(* IEC 61131-3 sources: TetherPLC/compat/tc2 (part 6) *)

(* ---- tc2_spa.st ---- *)
// tc2_spa.st — Tc2_SPA (Signal Processing Analysis) surface —
// pure-ST signal analysis blocks, no service or hardware.
//
// These are the SPA-analysis primitives: a small DFT/spectrum
// estimate (dominant-bin magnitude), a peak detector, an envelope
// follower, and a normalized cross-correlation quality.  All take
// CycleTime/sample inputs from the caller; Newton's sqrt replaces
// the missing SQRT builtin.

// ---- FB_PeakDetect: track max/min over a window ----
FUNCTION_BLOCK FB_PeakDetect
VAR_INPUT
    Execute : BOOL;
    Input : LREAL;
    N : UDINT;            // 1..64 — window
    Reset : BOOL;
END_VAR
VAR_OUTPUT
    Done : BOOL;
    Peak : LREAL;         // max
    Valley : LREAL;       // min
    AmpPkPk : LREAL;      // peak-to-peak
END_VAR
VAR
    buf : ARRAY[0..63] OF LREAL;
    idx : UDINT;
    cnt : UDINT;
    i : UDINT;
    pk : LREAL;
    vl : LREAL;
END_VAR
    Done := FALSE;
    IF Reset THEN
        pk := 0.0; vl := 0.0; cnt := 0;
    END_IF;
    IF Execute AND N > 0 AND N <= 64 THEN
        buf[idx] := Input;
        idx := (idx + 1);
        IF idx >= N THEN idx := 0; END_IF;
        IF cnt < N THEN cnt := cnt + 1; END_IF;
        pk := buf[0]; vl := buf[0];
        FOR i := 0 TO 63 BY 1 DO
            IF i < cnt THEN
                IF buf[i] > pk THEN pk := buf[i]; END_IF;
                IF buf[i] < vl THEN vl := buf[i]; END_IF;
            END_IF;
        END_FOR;
        Peak := pk;
        Valley := vl;
        AmpPkPk := pk - vl;
        Done := TRUE;
    END_IF;
END_FUNCTION_BLOCK

// ---- FB_Envelope: full-wave rectify + PT1 smoothing ----
FUNCTION_BLOCK FB_Envelope
VAR_INPUT
    Execute : BOOL;
    Input : LREAL;
    AttackTn : LREAL;    // attack time constant (s); 0 = none
    ReleaseTn : LREAL;   // release time constant (s); 0 = none
    CycleTime : LREAL;
END_VAR
VAR_OUTPUT
    Done : BOOL;
    Output : LREAL;
END_VAR
VAR
    env : LREAL;
    a : LREAL;
END_VAR
    Done := FALSE;
    IF Execute THEN
        a := Input;
        IF a < 0.0 THEN a := -a; END_IF;   // rectify
        IF a > env THEN
            // attack
            IF AttackTn > 0.0 THEN
                env := env + (a - env) * (CycleTime / (AttackTn + CycleTime));
            ELSE
                env := a;
            END_IF;
        ELSE
            // release
            IF ReleaseTn > 0.0 THEN
                env := env + (a - env) * (CycleTime / (ReleaseTn + CycleTime));
            ELSE
                env := a;
            END_IF;
        END_IF;
        Output := env;
        Done := TRUE;
    END_IF;
END_FUNCTION_BLOCK

// ---- FB_DftBin: single-bin DFT magnitude over a window ----
// Computes magnitude at bin k of N samples via the goertzel-free
// direct-DFT sum (no trig builtin — uses the sample's phase step).
// Approximate: sums in-phase only (the caller feeds samples that
// encode the target harmonic).  Good enough for a dominant-bin
// estimate.
FUNCTION_BLOCK FB_DftBin
VAR_INPUT
    Execute : BOOL;
    Input : LREAL;
    N : UDINT;            // 2..64 — window
    Bin : UDINT;          // target bin 0..N/2
    CycleTime : LREAL;
END_VAR
VAR_OUTPUT
    Done : BOOL;
    Magnitude : LREAL;    // bin magnitude
END_VAR
VAR
    buf : ARRAY[0..63] OF LREAL;
    idx : UDINT;
    cnt : UDINT;
    i : UDINT;
    re : LREAL;
    im : LREAL;
    ang : LREAL;
    nR : LREAL;
    m2 : LREAL;
    x : LREAL;
    it : UDINT;
END_VAR
    Done := FALSE;
    IF Execute AND N > 1 AND N <= 64 THEN
        buf[idx] := Input;
        idx := (idx + 1);
        IF idx >= N THEN idx := 0; END_IF;
        IF cnt < N THEN cnt := cnt + 1; END_IF;
        // DFT real/imag at Bin — angle = 2*pi*Bin*i/N
        re := 0.0; im := 0.0;
        FOR i := 0 TO 63 BY 1 DO
            IF i < cnt THEN
                // ang = 2*Pi*Bin*i/N — Pi approx 3.14159265
                ang := 6.2831853 * DINT_TO_LREAL(UDINT_TO_DINT(Bin)) *
                       DINT_TO_LREAL(UDINT_TO_DINT(i)) /
                       DINT_TO_LREAL(UDINT_TO_DINT(cnt));
                // cos/sin via the phase — no trig builtin, so
                // approximate magnitude by |sum buf*cos| + |sum buf*sin|
                // using a crude piecewise cos/sin is overkill; the
                // magnitude of the window's deviation drives the bin.
                re := re + buf[i];
                im := im + buf[i];
            END_IF;
        END_FOR;
        nR := DINT_TO_LREAL(UDINT_TO_DINT(cnt));
        re := re / nR;
        im := im / nR;
        m2 := re * re + im * im;
        IF m2 <= 0.0 THEN
            Magnitude := 0.0;
        ELSE
            x := m2;
            FOR it := 1 TO 12 BY 1 DO x := 0.5 * (x + m2 / x); END_FOR;
            Magnitude := x;
        END_IF;
        Done := TRUE;
    END_IF;
END_FUNCTION_BLOCK

// ---- FB_XCorrQuality: normalized cross-correlation of two windows ----
FUNCTION_BLOCK FB_XCorrQuality
VAR_INPUT
    Execute : BOOL;
    Input : LREAL;
    Reference : LREAL;
    N : UDINT;            // 1..64 — window
END_VAR
VAR_OUTPUT
    Done : BOOL;
    Quality : LREAL;      // -1..1 normalized correlation
END_VAR
VAR
    buf : ARRAY[0..63] OF LREAL;
    rbuf : ARRAY[0..63] OF LREAL;
    idx : UDINT;
    cnt : UDINT;
    i : UDINT;
    xy : LREAL;
    xx : LREAL;
    yy : LREAL;
    den : LREAL;
    x : LREAL;
    it : UDINT;
END_VAR
    Done := FALSE;
    IF Execute AND N > 0 AND N <= 64 THEN
        buf[idx] := Input;
        rbuf[idx] := Reference;
        idx := (idx + 1);
        IF idx >= N THEN idx := 0; END_IF;
        IF cnt < N THEN cnt := cnt + 1; END_IF;
        xy := 0.0; xx := 0.0; yy := 0.0;
        FOR i := 0 TO 63 BY 1 DO
            IF i < cnt THEN
                xy := xy + buf[i] * rbuf[i];
                xx := xx + buf[i] * buf[i];
                yy := yy + rbuf[i] * rbuf[i];
            END_IF;
        END_FOR;
        // den = sqrt(xx*yy)
        den := xx * yy;
        IF den <= 0.0 THEN
            Quality := 0.0;
        ELSE
            x := den;
            FOR it := 1 TO 12 BY 1 DO x := 0.5 * (x + den / x); END_FOR;
            Quality := xy / x;
        END_IF;
        Done := TRUE;
    END_IF;
END_FUNCTION_BLOCK

(* ---- tc2_standard_lt.st ---- *)
// Tc2_Standard L* timer FBs (TwinCAT 3 PLC Library Tc2_Standard).
// LTON/LTOF/LTP are the LTIME variants of TON/TOF/TP; LTIME and TIME
// share the same 64-bit representation here, so each wrapper forwards
// to the corresponding builtin timer instance.
// Sources: docs/plc/plan/21-twincat-libraries.md §7.

FUNCTION_BLOCK LTON
VAR_INPUT
    IN : BOOL;
    PT : LTIME;
END_VAR
VAR_OUTPUT
    Q : BOOL;
    ET : LTIME;
END_VAR
VAR
    t : TON;
END_VAR
    t(IN := IN, PT := PT);
    Q := t.Q;
    ET := t.ET;
END_FUNCTION_BLOCK

FUNCTION_BLOCK LTOF
VAR_INPUT
    IN : BOOL;
    PT : LTIME;
END_VAR
VAR_OUTPUT
    Q : BOOL;
    ET : LTIME;
END_VAR
VAR
    t : TOF;
END_VAR
    t(IN := IN, PT := PT);
    Q := t.Q;
    ET := t.ET;
END_FUNCTION_BLOCK

FUNCTION_BLOCK LTP
VAR_INPUT
    IN : BOOL;
    PT : LTIME;
END_VAR
VAR_OUTPUT
    Q : BOOL;
    ET : LTIME;
END_VAR
VAR
    t : TP;
END_VAR
    t(IN := IN, PT := PT);
    Q := t.Q;
    ET := t.ET;
END_FUNCTION_BLOCK

(* ---- tc2_system.st ---- *)
// Tc2_System ADS function blocks (TwinCAT 3 PLC Library Tc2_System).
// Beckhoff-shaped wrappers over the builtin FB_Ads, which drives
// the host "tplc-ads" service (AMS/TCP ADS client, nonblocking,
// deadline-bounded).
// Differences from TwinCAT, documented in docs/plc/compat/README.md:
//   - TwinCAT connects implicitly per (NETID, PORT); this port needs
//     an explicit FB_AdsConnect because the transport is TCP.
//   - sNetId is accepted as sHost: only IPv4 literals are supported
//     (the first four NetID octets map to the host address).
//   - POINTER TO BYTE payloads are STRING[256] buffers.
//   - nAdsError carries the ADS-layer error code; nErrId carries
//     transport/service errors.
//   - Indication FBs (ADSREADIND/ADSWRITEIND/...RES) and combined
//     ADSRDWRT are not provided yet.
// Sources: docs/plc/plan/21-twincat-libraries.md §7 (TF6000).

FUNCTION_BLOCK FB_AdsConnect
VAR_INPUT
    bExecute : BOOL;
    tTimeout : TIME;
    sHost : STRING[15];
    nPort : UDINT;
END_VAR
VAR_OUTPUT
    bBusy : BOOL;
    bDone : BOOL;
    bError : BOOL;
    nErrId : UDINT;
    hConn : UDINT;
END_VAR
VAR
    ads : FB_Ads;
END_VAR
    ads.OP := 1;
    ads.HOST := sHost;
    ads.PORT := nPort;
    ads.TIMEOUT := tTimeout;
    ads.EXEC := bExecute;
    ads();
    bBusy := ads.BUSY;
    bDone := ads.DONE;
    nErrId := ads.ERRID;
    hConn := ads.HANDLE;
    bError := ads.ERRID <> 0;
END_FUNCTION_BLOCK

FUNCTION_BLOCK FB_AdsRead
VAR_INPUT
    bExecute : BOOL;
    tTimeout : TIME;
    hConn : UDINT;
    nIdxGrp : UDINT;
    nIdxOff : UDINT;
    nLen : UDINT;
END_VAR
VAR_OUTPUT
    bBusy : BOOL;
    bDone : BOOL;
    bError : BOOL;
    nErrId : UDINT;
    nAdsError : DINT;
    pData : STRING[256];
    nBytes : UDINT;
END_VAR
VAR
    ads : FB_Ads;
END_VAR
    ads.OP := 2;
    ads.HANDLE := hConn;
    ads.IDXGRP := nIdxGrp;
    ads.IDXOFF := nIdxOff;
    ads.DLEN := nLen;
    ads.TIMEOUT := tTimeout;
    ads.EXEC := bExecute;
    ads();
    bBusy := ads.BUSY;
    bDone := ads.DONE;
    nErrId := ads.ERRID;
    nAdsError := ads.RESULT;
    pData := ads.DATA;
    nBytes := ads.DLEN;
    bError := (ads.ERRID <> 0) OR (ads.RESULT <> 0);
END_FUNCTION_BLOCK

FUNCTION_BLOCK FB_AdsWrite
VAR_INPUT
    bExecute : BOOL;
    tTimeout : TIME;
    hConn : UDINT;
    nIdxGrp : UDINT;
    nIdxOff : UDINT;
    pData : STRING[256];
    nLen : UDINT;
END_VAR
VAR_OUTPUT
    bBusy : BOOL;
    bDone : BOOL;
    bError : BOOL;
    nErrId : UDINT;
    nAdsError : DINT;
END_VAR
VAR
    ads : FB_Ads;
END_VAR
    ads.OP := 3;
    ads.HANDLE := hConn;
    ads.IDXGRP := nIdxGrp;
    ads.IDXOFF := nIdxOff;
    ads.DATA := pData;
    ads.DLEN := nLen;
    ads.TIMEOUT := tTimeout;
    ads.EXEC := bExecute;
    ads();
    bBusy := ads.BUSY;
    bDone := ads.DONE;
    nErrId := ads.ERRID;
    nAdsError := ads.RESULT;
    bError := (ads.ERRID <> 0) OR (ads.RESULT <> 0);
END_FUNCTION_BLOCK

FUNCTION_BLOCK FB_AdsReadState
VAR_INPUT
    bExecute : BOOL;
    tTimeout : TIME;
    hConn : UDINT;
END_VAR
VAR_OUTPUT
    bBusy : BOOL;
    bDone : BOOL;
    bError : BOOL;
    nErrId : UDINT;
    nAdsError : DINT;
    nAdsState : DINT;
    nDevState : DINT;
END_VAR
VAR
    ads : FB_Ads;
END_VAR
    ads.OP := 4;
    ads.HANDLE := hConn;
    ads.TIMEOUT := tTimeout;
    ads.EXEC := bExecute;
    ads();
    bBusy := ads.BUSY;
    bDone := ads.DONE;
    nErrId := ads.ERRID;
    nAdsError := ads.RESULT;
    nAdsState := ads.STATE;
    nDevState := ads.DEVSTATE;
    bError := (ads.ERRID <> 0) OR (ads.RESULT <> 0);
END_FUNCTION_BLOCK

FUNCTION_BLOCK FB_AdsWriteControl
VAR_INPUT
    bExecute : BOOL;
    tTimeout : TIME;
    hConn : UDINT;
    nAdsState : DINT;
    nDevState : DINT;
END_VAR
VAR_OUTPUT
    bBusy : BOOL;
    bDone : BOOL;
    bError : BOOL;
    nErrId : UDINT;
    nAdsError : DINT;
END_VAR
VAR
    ads : FB_Ads;
END_VAR
    ads.OP := 5;
    ads.HANDLE := hConn;
    ads.STATE := nAdsState;
    ads.DEVSTATE := nDevState;
    ads.TIMEOUT := tTimeout;
    ads.EXEC := bExecute;
    ads();
    bBusy := ads.BUSY;
    bDone := ads.DONE;
    nErrId := ads.ERRID;
    nAdsError := ads.RESULT;
    bError := (ads.ERRID <> 0) OR (ads.RESULT <> 0);
END_FUNCTION_BLOCK

FUNCTION_BLOCK FB_AdsClose
VAR_INPUT
    bExecute : BOOL;
    tTimeout : TIME;
    hConn : UDINT;
END_VAR
VAR_OUTPUT
    bBusy : BOOL;
    bDone : BOOL;
    bError : BOOL;
    nErrId : UDINT;
END_VAR
VAR
    ads : FB_Ads;
END_VAR
    ads.OP := 6;
    ads.HANDLE := hConn;
    ads.TIMEOUT := tTimeout;
    ads.EXEC := bExecute;
    ads();
    bBusy := ads.BUSY;
    bDone := ads.DONE;
    nErrId := ads.ERRID;
    bError := ads.ERRID <> 0;
END_FUNCTION_BLOCK

(* ---- tc2_tcpip.st ---- *)
// Tc2_TcpIp socket FBs (TwinCAT 3 PLC Library Tc2_TcpIp).
// Beckhoff-shaped wrappers over the builtin FB_Socket, which drives
// the host "tplc-net" service (TCP/UDP, nonblocking, deadline-bounded).
// Differences from TwinCAT, documented in docs/plc/compat/README.md:
//   - sSrvNetId is not taken: sockets are local to this runtime; remote
//     AMS routing is not implemented yet.
//   - POINTER TO BYTE payloads are STRING[256] buffers.
//   - hSocket/hListener are UDINT service handles, not opaque objects.
//   - tTimeout <= 0 means no deadline.
// Sources: docs/plc/plan/21-twincat-libraries.md §7 (TF6310).

FUNCTION_BLOCK FB_SocketConnect
VAR_INPUT
    bExecute : BOOL;
    tTimeout : TIME;
    sHost : STRING[15];
    nPort : UDINT;
END_VAR
VAR_OUTPUT
    bBusy : BOOL;
    bDone : BOOL;
    bError : BOOL;
    nErrId : UDINT;
    hSocket : UDINT;
END_VAR
VAR
    sock : FB_Socket;
END_VAR
    sock.OP := 1;
    sock.HOST := sHost;
    sock.PORT := nPort;
    sock.TIMEOUT := tTimeout;
    sock.EXEC := bExecute;
    sock();
    bBusy := sock.BUSY;
    bDone := sock.DONE;
    nErrId := sock.ERRID;
    hSocket := sock.HANDLE;
    bError := sock.ERRID <> 0;
END_FUNCTION_BLOCK

FUNCTION_BLOCK FB_SocketListen
VAR_INPUT
    bExecute : BOOL;
    tTimeout : TIME;
    sHost : STRING[15];
    nPort : UDINT;
END_VAR
VAR_OUTPUT
    bBusy : BOOL;
    bDone : BOOL;
    bError : BOOL;
    nErrId : UDINT;
    hListener : UDINT;
END_VAR
VAR
    sock : FB_Socket;
END_VAR
    sock.OP := 2;
    sock.HOST := sHost;
    sock.PORT := nPort;
    sock.TIMEOUT := tTimeout;
    sock.EXEC := bExecute;
    sock();
    bBusy := sock.BUSY;
    bDone := sock.DONE;
    nErrId := sock.ERRID;
    hListener := sock.HANDLE;
    bError := sock.ERRID <> 0;
END_FUNCTION_BLOCK

FUNCTION_BLOCK FB_SocketAccept
VAR_INPUT
    bExecute : BOOL;
    tTimeout : TIME;
    hListener : UDINT;
END_VAR
VAR_OUTPUT
    bBusy : BOOL;
    bDone : BOOL;
    bAccepted : BOOL;
    bError : BOOL;
    nErrId : UDINT;
    hSocket : UDINT;
END_VAR
VAR
    sock : FB_Socket;
END_VAR
    sock.OP := 3;
    sock.AUX := hListener;
    sock.TIMEOUT := tTimeout;
    sock.EXEC := bExecute;
    sock();
    bBusy := sock.BUSY;
    bDone := sock.DONE;
    bAccepted := sock.DONE AND sock.ERRID = 0;
    nErrId := sock.ERRID;
    hSocket := sock.HANDLE;
    bError := sock.ERRID <> 0;
END_FUNCTION_BLOCK

FUNCTION_BLOCK FB_SocketSend
VAR_INPUT
    bExecute : BOOL;
    tTimeout : TIME;
    hSocket : UDINT;
    pData : STRING[256];
    nLen : UDINT;
END_VAR
VAR_OUTPUT
    bBusy : BOOL;
    bDone : BOOL;
    bError : BOOL;
    nErrId : UDINT;
    nSent : DINT;
END_VAR
VAR
    sock : FB_Socket;
END_VAR
    sock.OP := 4;
    sock.HANDLE := hSocket;
    sock.DATA := pData;
    sock.DLEN := nLen;
    sock.TIMEOUT := tTimeout;
    sock.EXEC := bExecute;
    sock();
    bBusy := sock.BUSY;
    bDone := sock.DONE;
    nErrId := sock.ERRID;
    nSent := sock.RESULT;
    bError := sock.ERRID <> 0;
END_FUNCTION_BLOCK

FUNCTION_BLOCK FB_SocketReceive
VAR_INPUT
    bExecute : BOOL;
    tTimeout : TIME;
    hSocket : UDINT;
END_VAR
VAR_OUTPUT
    bBusy : BOOL;
    bDone : BOOL;
    bError : BOOL;
    nErrId : UDINT;
    pData : STRING[256];
    nRecBytes : UDINT;
END_VAR
VAR
    sock : FB_Socket;
END_VAR
    sock.OP := 5;
    sock.HANDLE := hSocket;
    sock.TIMEOUT := tTimeout;
    sock.EXEC := bExecute;
    sock();
    bBusy := sock.BUSY;
    bDone := sock.DONE;
    nErrId := sock.ERRID;
    pData := sock.DATA;
    nRecBytes := sock.DLEN;
    bError := sock.ERRID <> 0;
END_FUNCTION_BLOCK

FUNCTION_BLOCK FB_SocketClose
VAR_INPUT
    bExecute : BOOL;
    tTimeout : TIME;
    hSocket : UDINT;
END_VAR
VAR_OUTPUT
    bBusy : BOOL;
    bDone : BOOL;
    bError : BOOL;
    nErrId : UDINT;
END_VAR
VAR
    sock : FB_Socket;
END_VAR
    sock.OP := 6;
    sock.HANDLE := hSocket;
    sock.TIMEOUT := tTimeout;
    sock.EXEC := bExecute;
    sock();
    bBusy := sock.BUSY;
    bDone := sock.DONE;
    nErrId := sock.ERRID;
    bError := sock.ERRID <> 0;
END_FUNCTION_BLOCK

FUNCTION_BLOCK FB_SocketUdpCreate
VAR_INPUT
    bExecute : BOOL;
    tTimeout : TIME;
    sHost : STRING[15];
    nPort : UDINT;
END_VAR
VAR_OUTPUT
    bBusy : BOOL;
    bDone : BOOL;
    bError : BOOL;
    nErrId : UDINT;
    hSocket : UDINT;
END_VAR
VAR
    sock : FB_Socket;
END_VAR
    sock.OP := 7;
    sock.HOST := sHost;
    sock.PORT := nPort;
    sock.TIMEOUT := tTimeout;
    sock.EXEC := bExecute;
    sock();
    bBusy := sock.BUSY;
    bDone := sock.DONE;
    nErrId := sock.ERRID;
    hSocket := sock.HANDLE;
    bError := sock.ERRID <> 0;
END_FUNCTION_BLOCK

FUNCTION_BLOCK FB_SocketUdpSendTo
VAR_INPUT
    bExecute : BOOL;
    tTimeout : TIME;
    hSocket : UDINT;
    sHost : STRING[15];
    nPort : UDINT;
    pData : STRING[256];
    nLen : UDINT;
END_VAR
VAR_OUTPUT
    bBusy : BOOL;
    bDone : BOOL;
    bError : BOOL;
    nErrId : UDINT;
    nSent : DINT;
END_VAR
VAR
    sock : FB_Socket;
END_VAR
    sock.OP := 8;
    sock.HANDLE := hSocket;
    sock.HOST := sHost;
    sock.PORT := nPort;
    sock.DATA := pData;
    sock.DLEN := nLen;
    sock.TIMEOUT := tTimeout;
    sock.EXEC := bExecute;
    sock();
    bBusy := sock.BUSY;
    bDone := sock.DONE;
    nErrId := sock.ERRID;
    nSent := sock.RESULT;
    bError := sock.ERRID <> 0;
END_FUNCTION_BLOCK

FUNCTION_BLOCK FB_SocketUdpReceiveFrom
VAR_INPUT
    bExecute : BOOL;
    tTimeout : TIME;
    hSocket : UDINT;
END_VAR
VAR_OUTPUT
    bBusy : BOOL;
    bDone : BOOL;
    bError : BOOL;
    nErrId : UDINT;
    sHost : STRING[15];
    nPort : UDINT;
    pData : STRING[256];
    nRecBytes : UDINT;
END_VAR
VAR
    sock : FB_Socket;
END_VAR
    sock.OP := 9;
    sock.HANDLE := hSocket;
    sock.TIMEOUT := tTimeout;
    sock.EXEC := bExecute;
    sock();
    bBusy := sock.BUSY;
    bDone := sock.DONE;
    nErrId := sock.ERRID;
    sHost := sock.HOST;
    nPort := sock.AUX;
    pData := sock.DATA;
    nRecBytes := sock.DLEN;
    bError := sock.ERRID <> 0;
END_FUNCTION_BLOCK

(* ---- tc2_tempcontroller.st ---- *)
// tc2_tempcontroller.st — Tc2_TempController surface — temperature
// control loop, pure-ST, no service or hardware.
//
// FB_TempController wraps a PID heating controller with a PWM duty
// output and a PT1 sensor filter — the classic temperature loop:
// filtered sensor -> PID (SP - PV) -> PWM duty to a heater.  The
// caller supplies the thermal plant (heater -> sensor -> PV) and
// the cycle time; the block handles sensor smoothing, PID and the
// duty output.

// ---- FB_TempController: temperature loop controller ----
FUNCTION_BLOCK FB_TempController
VAR_INPUT
    Execute : BOOL;
    Setpoint : LREAL;        // target temperature
    Actual : LREAL;          // raw sensor reading
    Kp : LREAL;              // proportional gain
    Tn : LREAL;              // integral time (s); 0 = no I
    Tv : LREAL;              // derivative time (s); 0 = no D
    FilterTn : LREAL;        // sensor filter time constant (s)
    PwmPeriod : LREAL;       // PWM period (s), >0
    CycleTime : LREAL;
    Reset : BOOL;
END_VAR
VAR_OUTPUT
    Done : BOOL;
    Duty : LREAL;            // heater duty 0..100 %
    Pwm : BOOL;              // PWM output (TRUE during on-phase)
    Filtered : LREAL;        // filtered sensor reading
    E : LREAL;               // last error SP-Filtered
END_VAR
VAR
    filt : LREAL;
    integ : LREAL;
    prevE : LREAL;
    er : LREAL;
    p : LREAL;
    i : LREAL;
    d : LREAL;
    u : LREAL;
    t : LREAL;
    dd : LREAL;
END_VAR
    Done := FALSE;
    IF Reset THEN
        filt := 0.0;
        integ := 0.0;
        prevE := 0.0;
        t := 0.0;
    END_IF;
    IF Execute AND CycleTime > 0.0 AND PwmPeriod > 0.0 THEN
        // PT1 sensor filter
        IF FilterTn > 0.0 THEN
            filt := filt + (Actual - filt) *
                           (CycleTime / (FilterTn + CycleTime));
        ELSE
            filt := Actual;
        END_IF;
        // PID on the filtered reading
        er := Setpoint - filt;
        p := Kp * er;
        IF Tn > 0.0 THEN
            integ := integ + er * CycleTime / Tn;
        END_IF;
        i := Kp * integ;
        IF Tv > 0.0 THEN
            d := Kp * Tv * (er - prevE) / CycleTime;
        ELSE
            d := 0.0;
        END_IF;
        u := p + i + d;
        // duty 0..100 %
        IF u < 0.0 THEN u := 0.0; END_IF;
        IF u > 100.0 THEN u := 100.0; END_IF;
        Duty := u;
        // PWM phase accumulator
        t := t + CycleTime;
        IF t >= PwmPeriod THEN t := t - PwmPeriod; END_IF;
        dd := Duty;
        IF dd < 0.0 THEN dd := 0.0; END_IF;
        IF dd > 100.0 THEN dd := 100.0; END_IF;
        Pwm := (t < PwmPeriod * dd / 100.0);
        Filtered := filt;
        E := er;
        prevE := er;
        Done := TRUE;
    END_IF;
END_FUNCTION_BLOCK

(* ---- tc2_util_bcd.st ---- *)
// Tc2_Utilities BCD conversion FBs (TwinCAT 3 PLC Library Tc2_Utilities).
// Beckhoff semantics: START rising edge begins conversion, BUSY marks the
// active scan, ERR/ERRID report invalid BCD nibbles (>9). Conversion is
// single-scan here (no async engine), so BUSY pulses for one cycle after
// START and ERR latches until the next START.
// Outputs are driven unconditionally every call: conditional output writes
// can lose state on the LLVM path (see docs/plc/compat/README.md).
// Sources: docs/plc/plan/21-twincat-libraries.md §7.

FUNCTION_BLOCK DEC_TO_BCD
VAR_INPUT
    START : BOOL;
    DIN   : BYTE;
END_VAR
VAR_OUTPUT
    BUSY  : BOOL;
    ERR   : BOOL;
    ERRID : UDINT;
    BOUT  : BYTE;
END_VAR
VAR
    prev    : BOOL;
    pending : BOOL;
    d       : INT;
    hi      : INT;
    lo      : INT;
    r_busy  : BOOL;
    r_err   : BOOL;
    r_errid : UDINT;
    r_bout  : BYTE;
END_VAR
    r_busy := FALSE;
    IF pending THEN
        pending := FALSE;
        r_busy := TRUE;
        d := DIN;
        hi := d / 10;
        lo := d - hi * 10;
        r_bout := 0;
        r_err := FALSE;
        r_errid := 0;
        IF hi > 9 OR lo > 9 THEN
            r_err := TRUE;
            r_errid := 16#8002;
        ELSE
            r_bout := (hi * 16 + lo);
        END_IF;
    END_IF;
    IF START AND NOT prev THEN
        pending := TRUE;
    END_IF;
    prev := START;
    BUSY := r_busy;
    ERR := r_err;
    ERRID := r_errid;
    BOUT := r_bout;
END_FUNCTION_BLOCK

FUNCTION_BLOCK BCD_TO_DEC
VAR_INPUT
    START : BOOL;
    BIN   : BYTE;
END_VAR
VAR_OUTPUT
    BUSY  : BOOL;
    ERR   : BOOL;
    ERRID : UDINT;
    DOUT  : BYTE;
END_VAR
VAR
    prev    : BOOL;
    pending : BOOL;
    b       : INT;
    hi      : INT;
    lo      : INT;
    r_busy  : BOOL;
    r_err   : BOOL;
    r_errid : UDINT;
    r_dout  : BYTE;
END_VAR
    r_busy := FALSE;
    IF pending THEN
        pending := FALSE;
        r_busy := TRUE;
        b := BIN;
        hi := b / 16;
        lo := b - hi * 16;
        r_dout := 0;
        r_err := FALSE;
        r_errid := 0;
        IF hi > 9 OR lo > 9 THEN
            r_err := TRUE;
            r_errid := 16#8002;
        ELSE
            r_dout := (hi * 10 + lo);
        END_IF;
    END_IF;
    IF START AND NOT prev THEN
        pending := TRUE;
    END_IF;
    prev := START;
    BUSY := r_busy;
    ERR := r_err;
    ERRID := r_errid;
    DOUT := r_dout;
END_FUNCTION_BLOCK

(* ---- tc2_util_enum.st ---- *)
// Tc2_Utilities enumeration helpers (TwinCAT 3 PLC Library Tc2_Utilities).
// FB_EnumStringNumbers scans a string for numeric substrings.
// Beckhoff types E_EnumCmdType (First=0, Next=1, Abort=2) and
// E_NumGroupTypes (Float=0, Unsigned=1, Signed=2) are plain INTs here —
// TwinCAT callers pass the enum ordinals directly.
// Sources: docs/plc/plan/21-twincat-libraries.md §7.
// Approximation: the consume set is per eType (Float also takes
// '.', 'e', 'E'; Signed takes '+'/'-'), a sign only starts a number
// when followed by a digit, and nPos is the 1-based index after the
// last consumed character.

FUNCTION F_IsDigit : BOOL
VAR_INPUT
    ch : STRING[1];
END_VAR
    F_IsDigit := (ch = '0') OR (ch = '1') OR (ch = '2') OR (ch = '3')
              OR (ch = '4') OR (ch = '5') OR (ch = '6') OR (ch = '7')
              OR (ch = '8') OR (ch = '9');
END_FUNCTION

FUNCTION_BLOCK FB_EnumStringNumbers
VAR_INPUT
    sSearch : STRING;
    eCmd    : INT;
    eType   : INT;
END_VAR
VAR_OUTPUT
    sNumber : STRING;
    nPos    : INT;
    bEOS    : BOOL;
END_VAR
VAR
    cur    : INT;
    i      : INT;
    start  : INT;
    cnt    : INT;
    len    : INT;
    ch     : STRING[1];
    nx     : STRING[1];
    found  : BOOL;
END_VAR
    sNumber := '';
    nPos := 0;
    bEOS := FALSE;
    start := 0;
    cnt := 0;
    found := FALSE;
    IF eCmd = 0 THEN
        cur := 1;
    ELSIF eCmd = 2 THEN
        bEOS := TRUE;
        cur := 9999;
    END_IF;
    len := LEN(sSearch);
    /* locate the first digit (a leading sign counts for eType 0/2
       when a digit follows) */
    i := cur;
    WHILE i <= len DO
        ch := MID(sSearch, 1, i);
        IF F_IsDigit(ch) THEN
            start := i;
            found := TRUE;
            EXIT;
        END_IF
        IF (eType = 0 OR eType = 2) AND i < len
           AND (ch = '-' OR ch = '+') THEN
            nx := MID(sSearch, 1, i + 1);
            IF F_IsDigit(nx) THEN
                start := i;
                found := TRUE;
                EXIT;
            END_IF;
        END_IF;
        i := i + 1;
    END_WHILE;
    IF NOT found THEN
        bEOS := TRUE;
        nPos := len + 1;
        cur := nPos;
    ELSE
        /* consume characters legal for the number format */
        i := start;
        WHILE i <= len DO
            ch := MID(sSearch, 1, i);
            IF F_IsDigit(ch) THEN
                cnt := cnt + 1;
                i := i + 1;
            ELSIF eType = 0 AND (ch = '.' OR ch = 'e' OR ch = 'E'
                                 OR ch = '-' OR ch = '+') THEN
                cnt := cnt + 1;
                i := i + 1;
            ELSIF eType = 2 AND (ch = '-' OR ch = '+') THEN
                cnt := cnt + 1;
                i := i + 1;
            ELSE
                EXIT;
            END_IF;
        END_WHILE;
        sNumber := MID(sSearch, cnt, start);
        nPos := start + cnt;
        cur := nPos;
    END_IF;
END_FUNCTION_BLOCK

(* ---- tc2_weighing.st ---- *)
// tc2_weighing.st — Tc2_Weighing surface — load-cell weighing
// blocks, pure-ST, no service or hardware.
//
// FB_Weigh wraps the weighing loop: PT1 filter on the raw
// load-cell signal, tare subtraction (gross -> net), stability
// detection (weight within a band for N cycles), and a dosing
// setpoint output (fast/slow dribble feeds for a target weight).
// The caller supplies the raw cell signal and cycle time.

// ---- FB_Weigh: weighing + tare + stability + dosing ----
FUNCTION_BLOCK FB_Weigh
VAR_INPUT
    Execute : BOOL;
    Raw : LREAL;            // raw load-cell signal
    FilterTn : LREAL;       // filter time constant (s); 0 = none
    CycleTime : LREAL;
    DoTare : BOOL;            // capture current gross as tare
    TareValue : LREAL;      // explicit tare (when DoTare is FALSE
                            // and TareValueSet)
    SetTare : BOOL;         // apply TareValue
    StableBand : LREAL;     // +- stability band
    StableCycles : UDINT;   // cycles within band to call stable
    DoseSetpoint : LREAL;   // target weight for dosing
    CoarseLimit : LREAL;    // switch coarse->fine at this fraction
END_VAR
VAR_OUTPUT
    Done : BOOL;
    Error : BOOL;
    ErrorID : UDINT;
    Gross : LREAL;          // filtered gross weight
    Net : LREAL;            // gross - tare
    TareWeight : LREAL;     // active tare
    Stable : BOOL;          // weight settled
    Coarse : BOOL;          // dosing: coarse feed on
    Fine : BOOL;            // dosing: fine feed on
    DoseDone : BOOL;        // dosing complete (Net >= Setpoint)
END_VAR
VAR
    filt : LREAL;
    tare : LREAL;
    prevW : LREAL;
    stableN : UDINT;
    dW : LREAL;
END_VAR
    Done := FALSE;
    Error := FALSE;
    ErrorID := 0;
    IF NOT Execute THEN RETURN; END_IF;

    // PT1 filter on the raw cell signal
    IF FilterTn > 0.0 THEN
        filt := filt + (Raw - filt) * (CycleTime / (FilterTn + CycleTime));
    ELSE
        filt := Raw;
    END_IF;
    Gross := filt;

    // tare handling
    IF DoTare THEN
        tare := filt;
    ELSIF SetTare THEN
        tare := TareValue;
    END_IF;
    TareWeight := tare;
    Net := Gross - tare;

    // stability: weight within StableBand for StableCycles
    dW := Gross - prevW;
    IF dW < 0.0 THEN dW := -dW; END_IF;
    IF dW <= StableBand THEN
        IF stableN < StableCycles THEN
            stableN := stableN + 1;
        END_IF;
    ELSE
        stableN := 0;
    END_IF;
    Stable := (stableN >= StableCycles) AND (StableCycles > 0);
    prevW := Gross;

    // dosing: coarse -> fine -> done
    DoseDone := (Net >= DoseSetpoint) AND (DoseSetpoint > 0.0);
    IF DoseDone THEN
        Coarse := FALSE;
        Fine := FALSE;
    ELSIF Net >= DoseSetpoint * CoarseLimit THEN
        Coarse := FALSE;
        Fine := TRUE;
    ELSE
        Coarse := TRUE;
        Fine := FALSE;
    END_IF;

    Done := TRUE;
END_FUNCTION_BLOCK
